FUNCTION_BLOCK FB_IgorCtrl
VAR_INPUT
END_VAR
VAR_OUTPUT
	fbError:	FB_Error;
END_VAR
VAR
	fbPortal:			FB_Portal;
	fbSafetyMonitoring:	FB_SafetyMonitoring;
	fbFuseControl:		FB_FuseControl;
	fbFuseControl48V: 	FB_FuseControl_1;
	fbLight			:	FB_VI_Light;
END_VAR

VAR
	fbBlinkTimer1		: TON;
	fbBlinkTimer2		: TON;
	fbTimer				: TON;
	fbRS				: RS;
	nCntParty			: UINT;
	rTrig1				: R_TRIG;
	rTrig2				: R_TRIG;
	
	nRed				: UINT;
	nGreen				: UINT;
	nBlue				: UINT;
END_VAR

A_HmiComm();

fbSafetyMonitoring();

fbFuseControl();
fbFuseControl48V(bResetChannels := HMI.bQuit);


fbPortal(
	bFuseOk := NOT fbFuseControl.fbError.bError,
	bFuse48VOk := NOT fbFuseControl.fbError.bError,
	bManualMode:= HMI.bReqManualCtrl, 
	stNewJob:= HMI.stJob, 
	bImportJob:= HMI.bSetJob,
	bQuit:= HMI.bQuit OR fbPortal.bQuit,//kann quit nicht false setzen
	bSafetyRun := HMI.bSafetyRun,
	bSafetyOK=> HMI.bSafetyOK, 
	bBusy=> HMI.bPortalBusy,
	fbError=> );

HMI.bGripperClosed := fbPortal.fbGripper.bGripperClosed;
HMI.bGripperOpen := fbPortal.fbGripper.bGripperOpen;

IF NOT HMI.bSafetyRun AND NOT fbError.bError THEN
	fbError.M_Set(1, 'Steuerung ausgeschaltet', 0, E_ErrorIDs.eCtrlOff, E_ErrorSrcs.ePlc);
ELSIF HMI.bSafetyRun AND fbError.bError THEN
	fbError.M_Reset();
END_IF

//Set trigger white light
IF HMI.bLightOn THEN
	HMI.bLightWin := FALSE;
	HMI.bLightLose := FALSE;
	fbLight(bLightOn:= HMI.bLightOn);
	fbLight.bLightOn := FALSE;
	fbLight.SetIRGB(255, 255, 255, 255, 100);
ELSIF NOT HMI.bLightWin AND NOT HMI.bLightLose THEN
	fbLight(bLightOn:= HMI.bLightOn);
END_IF

//Set light for win
IF HMI.bLightWin AND NOT HMI.bLightLose AND NOT HMI.bLightOn THEN
	fbTimer(IN := TRUE, PT := T#3S);
	fbRS(SET := TRUE, RESET1 := fbTimer.Q);
	
	fbBlinkTimer1(IN := fbRS.Q1 AND NOT fbBlinkTimer2.Q, PT := T#0.5S, Q => fbLight.bLightOn);
	fbBlinkTimer2(IN := fbBlinkTimer1.Q, PT := T#0.5S);
	fbLight.SetIRGB(0, 0, 255, 0, 50);
	
	IF fbTimer.Q THEN
		HMI.bLightWin := FALSE;
		fbLight.bLightOn := FALSE;
		fbTimer(IN := FALSE);
		fbRS(SET := FALSE, RESET1 := TRUE);
	END_IF
	
	fbLight();
ELSE
	fbRS(SET := FALSE, RESET1 := FALSE);
END_IF

//set light for lose
IF HMI.bLightLose AND NOT HMI.bLightWin AND NOT HMI.bLightOn THEN
	fbTimer(IN := TRUE, PT := T#3S);
	fbRS(SET := TRUE, RESET1 := fbTimer.Q);
	
	fbBlinkTimer1(IN := fbRS.Q1 AND NOT fbBlinkTimer2.Q, PT := T#0.5S, Q => fbLight.bLightOn);
	fbBlinkTimer2(IN := fbBlinkTimer1.Q, PT := T#0.5S);
	fbLight.SetIRGB(0, 255, 0, 0, 50);
	
	IF fbTimer.Q THEN
		HMI.bLightLose := FALSE;
		fbLight.bLightOn := FALSE;
		fbTimer(IN := FALSE);
		fbRS(SET := FALSE, RESET1 := TRUE);
	END_IF
	
	fbLight();
ELSE
	fbRS(SET := FALSE, RESET1 := FALSE);
END_IF

//Party-Modus
IF HMI.bLightParty THEN
	fbTimer(IN := TRUE, PT := T#30S);
	fbRS(SET := TRUE, RESET1 := fbTimer.Q);
	
	fbBlinkTimer1(IN := fbRS.Q1 AND NOT fbBlinkTimer2.Q, PT := T#0.4S, Q => );
	fbBlinkTimer2(IN := fbBlinkTimer1.Q, PT := T#0.2S);
	fbLight.bLightOn := NOT fbBlinkTimer1.Q;
	IF rTrig1.Q OR rTrig2.Q THEN
		nCntParty := nCntParty + 1;
	END_IF
	
	CASE nCntParty OF 
		0: fbLight.SetIRGB(0, 255, 0, 0, 25);
		1: fbLight.SetIRGB(0, 255, 30, 0, 25);
		2: fbLight.SetIRGB(0, 255, 255, 0, 25);
		3: fbLight.SetIRGB(0, 180, 255, 0, 25);
		4: fbLight.SetIRGB(0, 0, 255, 0, 25);
		5: fbLight.SetIRGB(0, 0, 255, 150, 25);
		6: fbLight.SetIRGB(0, 0, 255, 255, 25);
		7: fbLight.SetIRGB(0, 0, 120, 255, 25);
		8: fbLight.SetIRGB(0, 0, 0, 255, 25);
		9: fbLight.SetIRGB(0, 120, 0, 255, 25);
		10: fbLight.SetIRGB(0, 255, 0, 120, 25); nCntParty := 0;
	END_CASE

	IF fbTimer.Q THEN
		HMI.bLightParty := FALSE;
		nCntParty := 0;
		fbLight.bLightOn := FALSE;
		fbTimer(IN := FALSE);
		fbRS(SET := FALSE, RESET1 := TRUE);
	END_IF
	
	rTrig1(CLK := fbBlinkTimer1.Q);
	rTrig2(CLK := fbBlinkTimer2.Q);
	fbLight();
ELSE
	fbRS(SET := FALSE, RESET1 := FALSE);
END_IF

ACTION A_HmiComm:
IF HMI.stSoftKeyCtrlOn.bIsPressed THEN
	HMI.bSafetyRun := TRUE;
END_IF
IF HMI.stSoftKeyCtrlOff.bIsPressed THEN
	HMI.bSafetyRun := FALSE;
END_IF
IF HMI.stSoftKeyAutoOn.bIsPressed THEN
	HMI.bReqManualCtrl := FALSE;
END_IF
IF HMI.stSoftKeyAutoOff.bIsPressed THEN
	HMI.bReqManualCtrl := TRUE;
END_IF

HMI.bInManual := MAIN.fbIgorCtrl.fbPortal.ePortalState = E_PortalState_New.eManualMode;

HMI.bHandInPortal := NOT MAIN.fbIgorCtrl.fbSafetyMonitoring.bLightCurtainOk;

HMI.bQuit := HMI.stSoftKeyQuit.bIsPressed;

IF HMI.bSafetyOK THEN
	HMI.stSoftKeyCtrlOn.eState := E_ButtonState_ON;
	HMI.stSoftKeyCtrlOff.eState := E_ButtonState_OFF;
	
	IF HMI.bReqManualCtrl THEN
		IF Main.fbIgorCtrl.fbPortal.ePortalState <> E_PortalState_New.eManualMode THEN
			HMI.stSoftKeyAutoOn.eState := E_ButtonState_BLINK;
			HMI.stSoftKeyAutoOff.eState := E_ButtonState_OFF;
		ELSE
			HMI.stSoftKeyAutoOn.eState := E_ButtonState_OFF;
			HMI.stSoftKeyAutoOff.eState := E_ButtonState_ON;
		END_IF
	ELSE
		IF HMI.nNumberErrors = 0 THEN
			HMI.stSoftKeyAutoOn.eState := E_ButtonState_ON;
			HMI.stSoftKeyAutoOff.eState := E_ButtonState_OFF;
		ELSE
			HMI.stSoftKeyAutoOn.eState := E_ButtonState_OFF;
			HMI.stSoftKeyAutoOff.eState := E_ButtonState_BLINK;
		END_IF
	END_IF
	
	IF HMI.nNumberErrors > 0 THEN
		HMI.stSoftKeyQuit.eState := E_ButtonState_BLINK;
	ELSE
		HMI.stSoftKeyQuit.eState := E_ButtonState_OFF;
	END_IF
ELSE
	HMI.stSoftKeyAutoOn.eState := E_ButtonState_OFF;
	HMI.stSoftKeyAutoOff.eState := E_ButtonState_ON;
	IF HMI.bSafetyRun THEN
		HMI.stSoftKeyCtrlOn.eState := E_ButtonState_BLINK;
		HMI.stSoftKeyCtrlOff.eState := E_ButtonState_OFF;
		HMI.stSoftKeyQuit.eState := E_ButtonState_BLINK;
	ELSE
		HMI.stSoftKeyCtrlOn.eState := E_ButtonState_OFF;
		HMI.stSoftKeyCtrlOff.eState := E_ButtonState_ON;
		HMI.stSoftKeyQuit.eState := E_ButtonState_OFF;
	END_IF
END_IF
END_ACTION

END_FUNCTION_BLOCK

(* stored: Version 1.1.0.1, ProductVersion 3.1.4024.12
   POU FB_IgorCtrl: Id {0fbc02e5-79f9-4bb2-a045-e538f92682ca}, SpecialFunc None
   Action A_HmiComm: Id {1d4a9ff5-a676-4205-9520-cd71c7a6778f} *)
